Yaskawa INFORM job: 20260625CHUFENGKOUFLIPOFFWELD.JBI

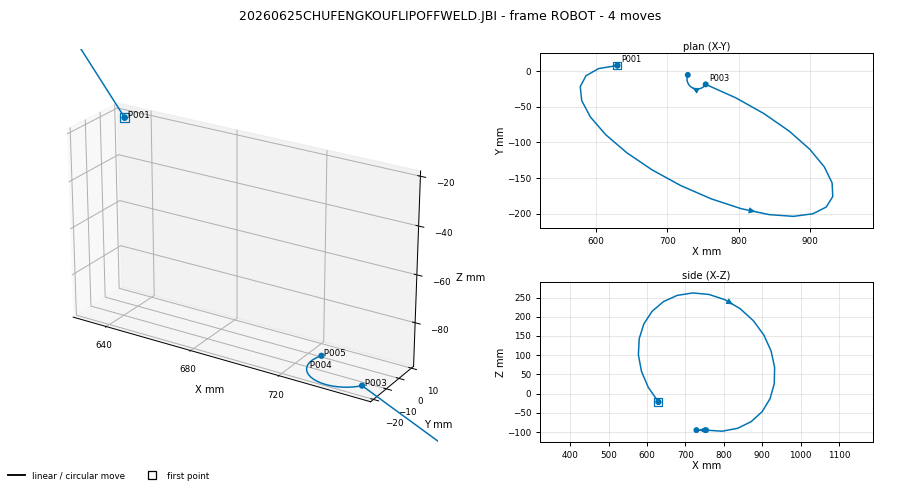
[picture p0: tool path of 20260625CHUFENGKOUFLIPOFFWELD.JBI in frame ROBOT, 4 of 9 moves have a stored position in this frame; points joined in program order, loops and branches not executed]
/JOB
//NAME 20260625CHUFENGKOUFLIPOFFWELD
//POS
///NPOS 3,0,3,5,0,5
///TOOL 1
///POSTYPE PULSE
///PULSE
C00000=-3653,-205,-30231,-2742,-71574,279
C00001=-3666,-425,-32327,-2755,-70295,311
C00002=-3332,9741,-5924,-2657,-80807,-35
///TOOL 0
EC00000=4,-321026
EC00001=4,-321026
EC00002=4,321023
///TOOL 1
///POSTYPE ROBOT
///RECTAN
///RCONF 0,0,0,0,0,0,0,0,0,0,0,0,0,0,0,0,0,0,0,0,0,0,0,0
P00001=629.883,8.042,-21.694,-154.9112,52.6025,29.7528
P00002=629.627,8.031,-21.395,-154.9194,52.6073,29.7435
P00003=753.895,-18.403,-95.100,179.0147,0.9881,-3.6266
P00004=729.189,-17.091,-95.012,179.5704,3.1491,-3.5911
P00005=728.757,-5.152,-95.055,179.5608,3.1535,-3.5736
///POSTYPE PULSE
///PULSE
EX00001=2,-321071
EX00002=2,321062
EX00003=0,0
EX00004=0,0
EX00005=0,0
//INST
///DATE 2026/06/25 14:50
///ATTR SC,RW
///GROUP1 RB1
///GROUP2 ST1
NOP
MOVJ C00000 VJ=0.78 PL=0  +MOVJ EC00000 VJ=0.78
MOVL C00001 V=11.0 PL=0  +MOVJ EC00001 VJ=0.78
MOVL P001 V=4.0 PL=0  +MOVJ EX001
SMOVC P001 V=4.0 PL=0  +MOVJ EX001
SMOVC P002 V=4.0 PL=0  +MOVJ EX002
SMOVC P003 V=4.0 PL=0  +MOVJ EX003
SMOVC P004 V=4.0 PL=0  +MOVJ EX004
SMOVC P005 V=4.0 PL=0  +MOVJ EX005
MOVL C00002 V=40.0 PL=0  +MOVJ EC00002 VJ=0.78
END
